TYPE ST_AxisControlResult :
STRUCT
Busy : BOOL;
Done : BOOL;
CommandAborted : BOOL;
Error : BOOL;
ErrorId : UDINT;
SourceErrorId : UDINT;
END_STRUCT
END_TYPE

(* stored: Version 1.1.0.1, ProductVersion 3.1.4026.20
   DUT ST_AxisControlResult: Id {6d61964b-e74e-5623-b41d-d027fabd9008} *)
